Fanuc KAREL source: KO00106.KL

PROGRAM KO00106
%NOLOCKGROUP
VAR
  A: REAL
  B: INTEGER
  OUT: REAL
BEGIN
  A = 1
  B = 2
  OUT = ATAN2(A, B)
END KO00106
